Fanuc KAREL source: KB00139.KL

PROGRAM KB00139
%NOLOCKGROUP
%ENVIRONMENT BYNAM
VAR
  P1: STRING[80]
  P2: INTEGER
  P3: INTEGER
  P4: INTEGER
  P5: ARRAY[4] OF STRING[80]
  P6: INTEGER
BEGIN
  P1 = 'A'
  P2 = 1
  P3 = 1
  P4 = 1
  P6 = 1
  PROG_LIST(P1, P2, P3, P4, P5, P6)
END KB00139
